(* IEC 61131-3 sources: PLC-Static-Analysis/modules/frontend-st/src/test/resources/dev/plca/frontend/st/StFrontendFuzzTestInputs/fuzzStText, 10 files *)

(* ---- types.st ---- *)
TYPE
    ST_Point EXTENDS ST_Base :
    STRUCT
        x : REAL;
        y : REAL := 0.0;
    END_STRUCT
    E_State : (Idle := 0, Running, Faulted := 10) INT := Idle;
    U_Raw :
    UNION
        dw : DWORD;
        ab : ARRAY[0..3] OF BYTE;
    END_UNION
    T_Name : STRING(80);
    T_Percent : INT(0..100);
    T_Matrix : ARRAY[1..3, 1..3] OF LREAL;
    T_Ref : REF_TO INT;
END_TYPE

(* ---- pragmas_comments.st ---- *)
// line comment
(* outer (* nested *) still outer *)
/* C-style /* nested */ comment */
{attribute 'qualified_only'}
{attribute 'TcLinkTo' := '.in := TIIB[Term 1]^Channel 1^Value'}
VAR_GLOBAL
    {attribute 'pytmc' := '
        pv: TEST:VALUE
        io: i
    '}
    gValue : INT; // trailing comment
    {warning 'check this'}
    gOther : INT;
END_VAR
{IF defined (SIMULATION)}
{ELSE}
{END_IF}
{region "Main part"}
{endregion}

(* ---- expressions.st ---- *)
FUNCTION F_Expr : LREAL
VAR_INPUT
    p : POINTER TO ST_Point;
END_VAR
VAR
    w : WORD;
    s : STRING;
    ws : WSTRING;
    b : BOOL;
    t : TIME;
END_VAR

F_Expr := -2 ** 2 + 3 * 4 MOD 5 - (1 + 2) / 3;
b := NOT b AND w.3 OR_ELSE p^.x > 1.5E-3 AND_THEN THIS^.bOk XOR SUPER^.bOk;
b := 1 < 2 = TRUE <> FALSE;
w := 16#FF_FF + 2#1010 + 8#17 + 10#99 + WORD#16#0F + INT#-5;
s := 'it$'s $N done';
ws := "wide $"quoted$"";
t := T#1h2m3s4ms + LTIME#-5us;
F_Expr := TO_LREAL(D#2024-01-31 - DATE#2024-01-01) + TOD#12:30:15.5 + DT#2024-01-31-12:00:00;
w := SIZEOF(POINTER TO ST_Point) + SIZEOF(STRING) + .gGlobal + AND(b, b);
F_Expr := arr[i, j + 1].field;
END_FUNCTION

(* ---- config_oop.st ---- *)
NAMESPACE Lib.Motion
USING Lib.Base, Other;
INTERFACE I_Axis EXTENDS I_Base, I_Diag
METHOD MoveAbs : BOOL
VAR_INPUT
    pos : LREAL;
END_VAR
END_METHOD
PROPERTY Position : LREAL
END_PROPERTY
END_INTERFACE
CLASS FINAL C_Axis IMPLEMENTS I_Axis
VAR PUBLIC
    pos : LREAL;
END_VAR
METHOD PUBLIC OVERRIDE MoveAbs : BOOL
MoveAbs := TRUE;
END_METHOD
END_CLASS
END_NAMESPACE

CONFIGURATION Cfg
VAR_GLOBAL
    gRun : BOOL;
END_VAR
RESOURCE Res ON PLC
    TASK Fast(INTERVAL := T#10MS, PRIORITY := 1);
    PROGRAM Main WITH Fast : MAIN;
END_RESOURCE
END_CONFIGURATION

(* ---- pou_function_block.st ---- *)
(* Function block with inheritance, all variable sections, methods, a property and an action. *)
{attribute 'reflection'}
FUNCTION_BLOCK PUBLIC FB_Motor EXTENDS FB_Base IMPLEMENTS I_Motor, I_Diag
VAR_INPUT
    bStart : BOOL;
    rSetpoint : REAL := 1.5;
END_VAR
VAR_OUTPUT
    bRunning AT %QX0.1 : BOOL;
END_VAR
VAR_IN_OUT
    stConfig : ST_Config;
END_VAR
VAR RETAIN PERSISTENT
    nStarts : UDINT;
END_VAR
VAR CONSTANT
    MAX_SPEED : INT := 1500;
END_VAR
VAR
    {attribute 'hide'}
    fbTimer : TON := (PT := T#2S);
    aBuf : ARRAY[0..9] OF INT := [1, 2, 8(0)];
    pData : POINTER TO BYTE;
    refCfg : REFERENCE TO ST_Config;
    fbInit : FB_Logger(10, sName := 'motor');
    a, b : INT;
END_VAR

fbTimer(IN := bStart, Q => bRunning);
IF bRunning THEN
    nStarts := nStarts + 1;
END_IF

METHOD PUBLIC Reset : BOOL
VAR_INPUT
    bForce : BOOL;
END_VAR
nStarts := 0;
Reset := TRUE;
END_METHOD

PROPERTY PUBLIC Speed : INT
GET
    Speed := MAX_SPEED;
END_GET
SET
    ;
END_SET
END_PROPERTY

ACTION Stop:
    bRunning := FALSE;
END_ACTION
END_FUNCTION_BLOCK

(* ---- text_export_no_end.st ---- *)
FUNCTION_BLOCK FB_Exported
VAR_INPUT
    bIn : BOOL;
END_VAR
VAR
    n : INT;
END_VAR
IF bIn THEN
    n := n + 1;
END_IF

(* ---- error_recovery.st ---- *)
PROGRAM P
VAR
    a : INT;
    b : INT := ;
    c : BOOL;
END_VAR
a := 1 +;
c := TRUE;
IF a > 1 THEN
    a := 2
END_IF
a FOO= 3;
§
c := FALSE;
b := 'unterminated
END_PROGRAM

(* ---- error_unterminated_comment.st ---- *)
PROGRAM P
VAR a : INT; END_VAR
a := 1;
(* this comment (* nests *) and is never closed
a := 2;

(* ---- statements.st ---- *)
PROGRAM MAIN
VAR
    i, n : INT;
    eState : E_State;
    bA, bB, bC : BOOL;
    r : REFERENCE TO INT;
    itf : I_Motor;
END_VAR

CASE eState OF
    E_State.Idle, E_State#Running:
        n := 1;
    1..5, 7:
        n := 2;
ELSE
    n := 0;
END_CASE;

FOR i := 0 TO 10 BY 2 DO
    IF i = 4 THEN CONTINUE; END_IF
    IF i > 8 THEN EXIT; END_IF
END_FOR

WHILE n < 10 DO n := n + 1; END_WHILE
REPEAT n := n - 1; UNTIL n <= 0 END_REPEAT

bA S= bB;
bA R= bC;
r REF= n;
itf ?= fbAny;
bA := bB := bC := FALSE;

JMP lbl;
lbl:
__TRY
    n := 1 / n;
__CATCH(exc)
    n := 0;
__FINALLY
    ;
__ENDTRY

fbT(IN := bA, PT := T#1S, Q => bB, NOT ET => );
RETURN;
END_PROGRAM

(* ---- statements_only.st ---- *)
// an exported action body: statements without any declaration
nCount := nCount + 1;
IF nCount > 10 THEN
    nCount := 0;
END_IF
